Fanuc KAREL source: KA00020.KL

PROGRAM KA00020
%NOLOCKGROUP
VAR
  SRC: REAL
  DST: JOINTPOS
BEGIN
  SRC = 2.0
  DST = SRC
END KA00020
